{attribute 'qualified_only'}
VAR_GLOBAL
  //---------------------------------------------------------------------------
  // MC2 encapsulation, CA movement
  //---------------------------------------------------------------------------
  MoverSelectorCtrl     : ST_MOVER_SELECTOR_CTRL;
  MoverSelectorState    : ST_MOVER_SELECTOR_STATE;
  //---------------------------------------------------------------------------
END_VAR

(* stored: Version 1.1.0.1
   GVL GVL_XTS: Id {09dfa152-1bd2-48eb-b928-a4a532d8b37f} *)
